Fanuc KAREL source: ko00033.KL

-- PROVISIONAL review KL for V770-1; original PC SHA256 9c486639ad807dbad0d3559372e1a4b050e3816f5d176554f8412119140c2df0
-- Incomplete behavior may be omitted. Consult companion uncertainty JSON. Do not deploy.
PROGRAM KO00033
%NOLOCKGROUP
BEGIN
  -- UNRESOLVED_PC offsets 5-12; opcodes 9D,23
  -- UNRESOLVED_PC offsets 17-66; opcodes 27,27,49,7E,AD,22,1C,22,31,7E,4A
  -- UNRESOLVED_PC offsets 71-75; opcodes 7F
END KO00033
